(* IEC 61131-3 sources: s7-to-codesys/tests/POUs/ScenariosLang/FB_BackwashGraph_ScenarioTest, 7 files *)

(* ---- FB_BackwashGraph_ScenarioTest.decl.st ---- *)
// AUTO-GENERATED — не редактировать: s7conv gen-tests, сценарии scenarios/lang/FB_BackwashGraph.csv
// Правка — в CSV (scenarios/README.md), затем python -m s7conv build-corpus.
// Назначение: тесты поведения сконвертированного FB_BackwashGraph по сценариям CSV (сценариев: 6, строк: 46):
//             один метод-тест на сценарий, строки — по порядку с моделируемым временем GVL_S7Clock.
//             Ожидаемые значения — из CSV (эталонные модели по описанию логики блока), не из
//             результата конвертации.
// Автор:      s7conv 0.1.0 (сгенерировано)
// Версия:     не указана
// Документ:   scenarios/README.md, docs/methodology.md, раздел «Проверка поведения»
FUNCTION_BLOCK FB_BackwashGraph_ScenarioTest EXTENDS coUnit.FB_TestSuite
VAR
    fbLongWash : FB_BackwashGraph;  // свой экземпляр на сценарий
    xLongWashDone : BOOL;  // сценарий выполнен (выполняется один раз)
    fbShortWash : FB_BackwashGraph;  // свой экземпляр на сценарий
    xShortWashDone : BOOL;  // сценарий выполнен (выполняется один раз)
    fbSupervision : FB_BackwashGraph;  // свой экземпляр на сценарий
    xSupervisionDone : BOOL;  // сценарий выполнен (выполняется один раз)
    fbAckSwitches : FB_BackwashGraph;  // свой экземпляр на сценарий
    xAckSwitchesDone : BOOL;  // сценарий выполнен (выполняется один раз)
    fbInterlockPump : FB_BackwashGraph;  // свой экземпляр на сценарий
    xInterlockPumpDone : BOOL;  // сценарий выполнен (выполняется один раз)
    fbOffAndInit : FB_BackwashGraph;  // свой экземпляр на сценарий
    xOffAndInitDone : BOOL;  // сценарий выполнен (выполняется один раз)
END_VAR

(* ---- AckSwitches.method.impl.st ---- *)
// AUTO-GENERATED — не редактировать: scenarios/lang/FB_BackwashGraph.csv, сценарий AckSwitches
coUnit.TEST('AckSwitches');
IF NOT xAckSwitchesDone THEN
    xAckSwitchesDone := TRUE;
    GVL_S7Clock.xSimulation := TRUE;

    // #1, t = 0 мс — первый вызов: начальный шаг Idle
    GVL_S7Clock.tSimNow := T#0MS;
    fbAckSwitches.OFF_SQ := FALSE;
    fbAckSwitches.INIT_SQ := FALSE;
    fbAckSwitches.ACK_EF := FALSE;
    fbAckSwitches.xStart := FALSE;
    fbAckSwitches.xLevelLow := FALSE;
    fbAckSwitches.xLevelHigh := FALSE;
    fbAckSwitches.xShortWash := FALSE;
    fbAckSwitches.xPumpOk := TRUE;
    fbAckSwitches.xValveFault := FALSE;
    fbAckSwitches();
    AssertEquals_BOOL(Expected := FALSE, Actual := fbAckSwitches.ERR_FLT, Message := 'AckSwitches#1 ERR_FLT');
    AssertEquals_BOOL(Expected := TRUE, Actual := fbAckSwitches.xReady, Message := 'AckSwitches#1 xReady');
    AssertEquals_BOOL(Expected := FALSE, Actual := fbAckSwitches.xDrainValve, Message := 'AckSwitches#1 xDrainValve');
    AssertEquals_BOOL(Expected := FALSE, Actual := fbAckSwitches.xBlower, Message := 'AckSwitches#1 xBlower');
    AssertEquals_BOOL(Expected := FALSE, Actual := fbAckSwitches.xAirValve, Message := 'AckSwitches#1 xAirValve');
    AssertEquals_BOOL(Expected := FALSE, Actual := fbAckSwitches.xWashPump, Message := 'AckSwitches#1 xWashPump');
    AssertEquals_BOOL(Expected := FALSE, Actual := fbAckSwitches.xInletValve, Message := 'AckSwitches#1 xInletValve');
    AssertEquals_BOOL(Expected := FALSE, Actual := fbAckSwitches.xWashActive, Message := 'AckSwitches#1 xWashActive');
    AssertEquals_BOOL(Expected := FALSE, Actual := fbAckSwitches.xValvesBusy, Message := 'AckSwitches#1 xValvesBusy');
    AssertEquals_INT(Expected := 0, Actual := fbAckSwitches.iWashCount, Message := 'AckSwitches#1 iWashCount');

    // #2, t = 100 мс — T1 Start: Drain, промывка №1, слив открыт
    GVL_S7Clock.tSimNow := T#100MS;
    fbAckSwitches.xStart := TRUE;
    fbAckSwitches();
    AssertEquals_BOOL(Expected := FALSE, Actual := fbAckSwitches.ERR_FLT, Message := 'AckSwitches#2 ERR_FLT');
    AssertEquals_BOOL(Expected := FALSE, Actual := fbAckSwitches.xReady, Message := 'AckSwitches#2 xReady');
    AssertEquals_BOOL(Expected := TRUE, Actual := fbAckSwitches.xDrainValve, Message := 'AckSwitches#2 xDrainValve');
    AssertEquals_BOOL(Expected := FALSE, Actual := fbAckSwitches.xBlower, Message := 'AckSwitches#2 xBlower');
    AssertEquals_BOOL(Expected := FALSE, Actual := fbAckSwitches.xAirValve, Message := 'AckSwitches#2 xAirValve');
    AssertEquals_BOOL(Expected := FALSE, Actual := fbAckSwitches.xWashPump, Message := 'AckSwitches#2 xWashPump');
    AssertEquals_BOOL(Expected := FALSE, Actual := fbAckSwitches.xInletValve, Message := 'AckSwitches#2 xInletValve');
    AssertEquals_BOOL(Expected := TRUE, Actual := fbAckSwitches.xWashActive, Message := 'AckSwitches#2 xWashActive');
    AssertEquals_BOOL(Expected := TRUE, Actual := fbAckSwitches.xValvesBusy, Message := 'AckSwitches#2 xValvesBusy');
    AssertEquals_INT(Expected := 1, Actual := fbAckSwitches.iWashCount, Message := 'AckSwitches#2 iWashCount');

    // #3, t = 200 мс — слив
    GVL_S7Clock.tSimNow := T#200MS;
    fbAckSwitches.xStart := FALSE;
    fbAckSwitches();
    AssertEquals_BOOL(Expected := FALSE, Actual := fbAckSwitches.ERR_FLT, Message := 'AckSwitches#3 ERR_FLT');
    AssertEquals_BOOL(Expected := FALSE, Actual := fbAckSwitches.xReady, Message := 'AckSwitches#3 xReady');
    AssertEquals_BOOL(Expected := TRUE, Actual := fbAckSwitches.xDrainValve, Message := 'AckSwitches#3 xDrainValve');
    AssertEquals_BOOL(Expected := FALSE, Actual := fbAckSwitches.xBlower, Message := 'AckSwitches#3 xBlower');
    AssertEquals_BOOL(Expected := FALSE, Actual := fbAckSwitches.xAirValve, Message := 'AckSwitches#3 xAirValve');
    AssertEquals_BOOL(Expected := FALSE, Actual := fbAckSwitches.xWashPump, Message := 'AckSwitches#3 xWashPump');
    AssertEquals_BOOL(Expected := FALSE, Actual := fbAckSwitches.xInletValve, Message := 'AckSwitches#3 xInletValve');
    AssertEquals_BOOL(Expected := TRUE, Actual := fbAckSwitches.xWashActive, Message := 'AckSwitches#3 xWashActive');
    AssertEquals_BOOL(Expected := TRUE, Actual := fbAckSwitches.xValvesBusy, Message := 'AckSwitches#3 xValvesBusy');
    AssertEquals_INT(Expected := 1, Actual := fbAckSwitches.iWashCount, Message := 'AckSwitches#3 iWashCount');

    // #4, t = 500 мс — ошибка контроля
    GVL_S7Clock.tSimNow := T#500MS;
    fbAckSwitches.xShortWash := TRUE;
    fbAckSwitches.xValveFault := TRUE;
    fbAckSwitches();
    AssertEquals_BOOL(Expected := TRUE, Actual := fbAckSwitches.ERR_FLT, Message := 'AckSwitches#4 ERR_FLT');
    AssertEquals_BOOL(Expected := FALSE, Actual := fbAckSwitches.xReady, Message := 'AckSwitches#4 xReady');
    AssertEquals_BOOL(Expected := TRUE, Actual := fbAckSwitches.xDrainValve, Message := 'AckSwitches#4 xDrainValve');
    AssertEquals_BOOL(Expected := FALSE, Actual := fbAckSwitches.xBlower, Message := 'AckSwitches#4 xBlower');
    AssertEquals_BOOL(Expected := FALSE, Actual := fbAckSwitches.xAirValve, Message := 'AckSwitches#4 xAirValve');
    AssertEquals_BOOL(Expected := FALSE, Actual := fbAckSwitches.xWashPump, Message := 'AckSwitches#4 xWashPump');
    AssertEquals_BOOL(Expected := FALSE, Actual := fbAckSwitches.xInletValve, Message := 'AckSwitches#4 xInletValve');
    AssertEquals_BOOL(Expected := TRUE, Actual := fbAckSwitches.xWashActive, Message := 'AckSwitches#4 xWashActive');
    AssertEquals_BOOL(Expected := TRUE, Actual := fbAckSwitches.xValvesBusy, Message := 'AckSwitches#4 xValvesBusy');
    AssertEquals_INT(Expected := 1, Actual := fbAckSwitches.iWashCount, Message := 'AckSwitches#4 iWashCount');

    // #5, t = 600 мс — квитирование и уровень: T3 ShortWash в том же вызове
    GVL_S7Clock.tSimNow := T#600MS;
    fbAckSwitches.ACK_EF := TRUE;
    fbAckSwitches.xLevelLow := TRUE;
    fbAckSwitches();
    AssertEquals_BOOL(Expected := FALSE, Actual := fbAckSwitches.ERR_FLT, Message := 'AckSwitches#5 ERR_FLT');
    AssertEquals_BOOL(Expected := FALSE, Actual := fbAckSwitches.xReady, Message := 'AckSwitches#5 xReady');
    AssertEquals_BOOL(Expected := FALSE, Actual := fbAckSwitches.xDrainValve, Message := 'AckSwitches#5 xDrainValve');
    AssertEquals_BOOL(Expected := FALSE, Actual := fbAckSwitches.xBlower, Message := 'AckSwitches#5 xBlower');
    AssertEquals_BOOL(Expected := FALSE, Actual := fbAckSwitches.xAirValve, Message := 'AckSwitches#5 xAirValve');
    AssertEquals_BOOL(Expected := TRUE, Actual := fbAckSwitches.xWashPump, Message := 'AckSwitches#5 xWashPump');
    AssertEquals_BOOL(Expected := FALSE, Actual := fbAckSwitches.xInletValve, Message := 'AckSwitches#5 xInletValve');
    AssertEquals_BOOL(Expected := TRUE, Actual := fbAckSwitches.xWashActive, Message := 'AckSwitches#5 xWashActive');
    AssertEquals_BOOL(Expected := FALSE, Actual := fbAckSwitches.xValvesBusy, Message := 'AckSwitches#5 xValvesBusy');
    AssertEquals_INT(Expected := 1, Actual := fbAckSwitches.iWashCount, Message := 'AckSwitches#5 iWashCount');

    // #6, t = 700 мс — QuickRinse: контроль Drain больше не действует
    GVL_S7Clock.tSimNow := T#700MS;
    fbAckSwitches.ACK_EF := FALSE;
    fbAckSwitches.xLevelLow := FALSE;
    fbAckSwitches();
    AssertEquals_BOOL(Expected := FALSE, Actual := fbAckSwitches.ERR_FLT, Message := 'AckSwitches#6 ERR_FLT');
    AssertEquals_BOOL(Expected := FALSE, Actual := fbAckSwitches.xReady, Message := 'AckSwitches#6 xReady');
    AssertEquals_BOOL(Expected := FALSE, Actual := fbAckSwitches.xDrainValve, Message := 'AckSwitches#6 xDrainValve');
    AssertEquals_BOOL(Expected := FALSE, Actual := fbAckSwitches.xBlower, Message := 'AckSwitches#6 xBlower');
    AssertEquals_BOOL(Expected := FALSE, Actual := fbAckSwitches.xAirValve, Message := 'AckSwitches#6 xAirValve');
    AssertEquals_BOOL(Expected := TRUE, Actual := fbAckSwitches.xWashPump, Message := 'AckSwitches#6 xWashPump');
    AssertEquals_BOOL(Expected := FALSE, Actual := fbAckSwitches.xInletValve, Message := 'AckSwitches#6 xInletValve');
    AssertEquals_BOOL(Expected := TRUE, Actual := fbAckSwitches.xWashActive, Message := 'AckSwitches#6 xWashActive');
    AssertEquals_BOOL(Expected := FALSE, Actual := fbAckSwitches.xValvesBusy, Message := 'AckSwitches#6 xValvesBusy');
    AssertEquals_INT(Expected := 1, Actual := fbAckSwitches.iWashCount, Message := 'AckSwitches#6 iWashCount');

    GVL_S7Clock.xSimulation := FALSE;
END_IF
coUnit.TEST_FINISHED();

(* ---- InterlockPump.method.impl.st ---- *)
// AUTO-GENERATED — не редактировать: scenarios/lang/FB_BackwashGraph.csv, сценарий InterlockPump
coUnit.TEST('InterlockPump');
IF NOT xInterlockPumpDone THEN
    xInterlockPumpDone := TRUE;
    GVL_S7Clock.xSimulation := TRUE;

    // #1, t = 0 мс — первый вызов: начальный шаг Idle
    GVL_S7Clock.tSimNow := T#0MS;
    fbInterlockPump.OFF_SQ := FALSE;
    fbInterlockPump.INIT_SQ := FALSE;
    fbInterlockPump.ACK_EF := FALSE;
    fbInterlockPump.xStart := FALSE;
    fbInterlockPump.xLevelLow := FALSE;
    fbInterlockPump.xLevelHigh := FALSE;
    fbInterlockPump.xShortWash := FALSE;
    fbInterlockPump.xPumpOk := TRUE;
    fbInterlockPump.xValveFault := FALSE;
    fbInterlockPump();
    AssertEquals_BOOL(Expected := FALSE, Actual := fbInterlockPump.ERR_FLT, Message := 'InterlockPump#1 ERR_FLT');
    AssertEquals_BOOL(Expected := TRUE, Actual := fbInterlockPump.xReady, Message := 'InterlockPump#1 xReady');
    AssertEquals_BOOL(Expected := FALSE,
                      Actual := fbInterlockPump.xDrainValve,
                      Message := 'InterlockPump#1 xDrainValve');
    AssertEquals_BOOL(Expected := FALSE, Actual := fbInterlockPump.xBlower, Message := 'InterlockPump#1 xBlower');
    AssertEquals_BOOL(Expected := FALSE, Actual := fbInterlockPump.xAirValve, Message := 'InterlockPump#1 xAirValve');
    AssertEquals_BOOL(Expected := FALSE, Actual := fbInterlockPump.xWashPump, Message := 'InterlockPump#1 xWashPump');
    AssertEquals_BOOL(Expected := FALSE,
                      Actual := fbInterlockPump.xInletValve,
                      Message := 'InterlockPump#1 xInletValve');
    AssertEquals_BOOL(Expected := FALSE,
                      Actual := fbInterlockPump.xWashActive,
                      Message := 'InterlockPump#1 xWashActive');
    AssertEquals_BOOL(Expected := FALSE,
                      Actual := fbInterlockPump.xValvesBusy,
                      Message := 'InterlockPump#1 xValvesBusy');
    AssertEquals_INT(Expected := 0, Actual := fbInterlockPump.iWashCount, Message := 'InterlockPump#1 iWashCount');

    // #2, t = 100 мс — T1 Start: Drain, промывка №1, слив открыт
    GVL_S7Clock.tSimNow := T#100MS;
    fbInterlockPump.xStart := TRUE;
    fbInterlockPump();
    AssertEquals_BOOL(Expected := FALSE, Actual := fbInterlockPump.ERR_FLT, Message := 'InterlockPump#2 ERR_FLT');
    AssertEquals_BOOL(Expected := FALSE, Actual := fbInterlockPump.xReady, Message := 'InterlockPump#2 xReady');
    AssertEquals_BOOL(Expected := TRUE,
                      Actual := fbInterlockPump.xDrainValve,
                      Message := 'InterlockPump#2 xDrainValve');
    AssertEquals_BOOL(Expected := FALSE, Actual := fbInterlockPump.xBlower, Message := 'InterlockPump#2 xBlower');
    AssertEquals_BOOL(Expected := FALSE, Actual := fbInterlockPump.xAirValve, Message := 'InterlockPump#2 xAirValve');
    AssertEquals_BOOL(Expected := FALSE, Actual := fbInterlockPump.xWashPump, Message := 'InterlockPump#2 xWashPump');
    AssertEquals_BOOL(Expected := FALSE,
                      Actual := fbInterlockPump.xInletValve,
                      Message := 'InterlockPump#2 xInletValve');
    AssertEquals_BOOL(Expected := TRUE,
                      Actual := fbInterlockPump.xWashActive,
                      Message := 'InterlockPump#2 xWashActive');
    AssertEquals_BOOL(Expected := TRUE,
                      Actual := fbInterlockPump.xValvesBusy,
                      Message := 'InterlockPump#2 xValvesBusy');
    AssertEquals_INT(Expected := 1, Actual := fbInterlockPump.iWashCount, Message := 'InterlockPump#2 iWashCount');

    // #3, t = 200 мс — слив
    GVL_S7Clock.tSimNow := T#200MS;
    fbInterlockPump.xStart := FALSE;
    fbInterlockPump();
    AssertEquals_BOOL(Expected := FALSE, Actual := fbInterlockPump.ERR_FLT, Message := 'InterlockPump#3 ERR_FLT');
    AssertEquals_BOOL(Expected := FALSE, Actual := fbInterlockPump.xReady, Message := 'InterlockPump#3 xReady');
    AssertEquals_BOOL(Expected := TRUE,
                      Actual := fbInterlockPump.xDrainValve,
                      Message := 'InterlockPump#3 xDrainValve');
    AssertEquals_BOOL(Expected := FALSE, Actual := fbInterlockPump.xBlower, Message := 'InterlockPump#3 xBlower');
    AssertEquals_BOOL(Expected := FALSE, Actual := fbInterlockPump.xAirValve, Message := 'InterlockPump#3 xAirValve');
    AssertEquals_BOOL(Expected := FALSE, Actual := fbInterlockPump.xWashPump, Message := 'InterlockPump#3 xWashPump');
    AssertEquals_BOOL(Expected := FALSE,
                      Actual := fbInterlockPump.xInletValve,
                      Message := 'InterlockPump#3 xInletValve');
    AssertEquals_BOOL(Expected := TRUE,
                      Actual := fbInterlockPump.xWashActive,
                      Message := 'InterlockPump#3 xWashActive');
    AssertEquals_BOOL(Expected := TRUE,
                      Actual := fbInterlockPump.xValvesBusy,
                      Message := 'InterlockPump#3 xValvesBusy');
    AssertEquals_INT(Expected := 1, Actual := fbInterlockPump.iWashCount, Message := 'InterlockPump#3 iWashCount');

    // #4, t = 1000 мс — Air и Rinse: насос промывки включён
    GVL_S7Clock.tSimNow := T#1000MS;
    fbInterlockPump.xLevelLow := TRUE;
    fbInterlockPump();
    AssertEquals_BOOL(Expected := FALSE, Actual := fbInterlockPump.ERR_FLT, Message := 'InterlockPump#4 ERR_FLT');
    AssertEquals_BOOL(Expected := FALSE, Actual := fbInterlockPump.xReady, Message := 'InterlockPump#4 xReady');
    AssertEquals_BOOL(Expected := FALSE,
                      Actual := fbInterlockPump.xDrainValve,
                      Message := 'InterlockPump#4 xDrainValve');
    AssertEquals_BOOL(Expected := TRUE, Actual := fbInterlockPump.xBlower, Message := 'InterlockPump#4 xBlower');
    AssertEquals_BOOL(Expected := FALSE, Actual := fbInterlockPump.xAirValve, Message := 'InterlockPump#4 xAirValve');
    AssertEquals_BOOL(Expected := TRUE, Actual := fbInterlockPump.xWashPump, Message := 'InterlockPump#4 xWashPump');
    AssertEquals_BOOL(Expected := FALSE,
                      Actual := fbInterlockPump.xInletValve,
                      Message := 'InterlockPump#4 xInletValve');
    AssertEquals_BOOL(Expected := TRUE,
                      Actual := fbInterlockPump.xWashActive,
                      Message := 'InterlockPump#4 xWashActive');
    AssertEquals_BOOL(Expected := FALSE,
                      Actual := fbInterlockPump.xValvesBusy,
                      Message := 'InterlockPump#4 xValvesBusy');
    AssertEquals_INT(Expected := 1, Actual := fbInterlockPump.iWashCount, Message := 'InterlockPump#4 iWashCount');

    // #5, t = 1100 мс — насос неисправен: блокировка не выполнена
    GVL_S7Clock.tSimNow := T#1100MS;
    fbInterlockPump.xLevelLow := FALSE;
    fbInterlockPump.xPumpOk := FALSE;
    fbInterlockPump();
    AssertEquals_BOOL(Expected := FALSE, Actual := fbInterlockPump.ERR_FLT, Message := 'InterlockPump#5 ERR_FLT');
    AssertEquals_BOOL(Expected := FALSE, Actual := fbInterlockPump.xReady, Message := 'InterlockPump#5 xReady');
    AssertEquals_BOOL(Expected := FALSE,
                      Actual := fbInterlockPump.xDrainValve,
                      Message := 'InterlockPump#5 xDrainValve');
    AssertEquals_BOOL(Expected := TRUE, Actual := fbInterlockPump.xBlower, Message := 'InterlockPump#5 xBlower');
    AssertEquals_BOOL(Expected := FALSE, Actual := fbInterlockPump.xAirValve, Message := 'InterlockPump#5 xAirValve');
    AssertEquals_BOOL(Expected := FALSE, Actual := fbInterlockPump.xWashPump, Message := 'InterlockPump#5 xWashPump');
    AssertEquals_BOOL(Expected := FALSE,
                      Actual := fbInterlockPump.xInletValve,
                      Message := 'InterlockPump#5 xInletValve');
    AssertEquals_BOOL(Expected := TRUE,
                      Actual := fbInterlockPump.xWashActive,
                      Message := 'InterlockPump#5 xWashActive');
    AssertEquals_BOOL(Expected := FALSE,
                      Actual := fbInterlockPump.xValvesBusy,
                      Message := 'InterlockPump#5 xValvesBusy');
    AssertEquals_INT(Expected := 1, Actual := fbInterlockPump.iWashCount, Message := 'InterlockPump#5 iWashCount');

    // #6, t = 1200 мс — насос исправен: снова включён
    GVL_S7Clock.tSimNow := T#1200MS;
    fbInterlockPump.xPumpOk := TRUE;
    fbInterlockPump();
    AssertEquals_BOOL(Expected := FALSE, Actual := fbInterlockPump.ERR_FLT, Message := 'InterlockPump#6 ERR_FLT');
    AssertEquals_BOOL(Expected := FALSE, Actual := fbInterlockPump.xReady, Message := 'InterlockPump#6 xReady');
    AssertEquals_BOOL(Expected := FALSE,
                      Actual := fbInterlockPump.xDrainValve,
                      Message := 'InterlockPump#6 xDrainValve');
    AssertEquals_BOOL(Expected := TRUE, Actual := fbInterlockPump.xBlower, Message := 'InterlockPump#6 xBlower');
    AssertEquals_BOOL(Expected := FALSE, Actual := fbInterlockPump.xAirValve, Message := 'InterlockPump#6 xAirValve');
    AssertEquals_BOOL(Expected := TRUE, Actual := fbInterlockPump.xWashPump, Message := 'InterlockPump#6 xWashPump');
    AssertEquals_BOOL(Expected := FALSE,
                      Actual := fbInterlockPump.xInletValve,
                      Message := 'InterlockPump#6 xInletValve');
    AssertEquals_BOOL(Expected := TRUE,
                      Actual := fbInterlockPump.xWashActive,
                      Message := 'InterlockPump#6 xWashActive');
    AssertEquals_BOOL(Expected := FALSE,
                      Actual := fbInterlockPump.xValvesBusy,
                      Message := 'InterlockPump#6 xValvesBusy');
    AssertEquals_INT(Expected := 1, Actual := fbInterlockPump.iWashCount, Message := 'InterlockPump#6 iWashCount');

    GVL_S7Clock.xSimulation := FALSE;
END_IF
coUnit.TEST_FINISHED();

(* ---- LongWash.method.impl.st ---- *)
// AUTO-GENERATED — не редактировать: scenarios/lang/FB_BackwashGraph.csv, сценарий LongWash
coUnit.TEST('LongWash');
IF NOT xLongWashDone THEN
    xLongWashDone := TRUE;
    GVL_S7Clock.xSimulation := TRUE;

    // #1, t = 0 мс — первый вызов: начальный шаг Idle
    GVL_S7Clock.tSimNow := T#0MS;
    fbLongWash.OFF_SQ := FALSE;
    fbLongWash.INIT_SQ := FALSE;
    fbLongWash.ACK_EF := FALSE;
    fbLongWash.xStart := FALSE;
    fbLongWash.xLevelLow := FALSE;
    fbLongWash.xLevelHigh := FALSE;
    fbLongWash.xShortWash := FALSE;
    fbLongWash.xPumpOk := TRUE;
    fbLongWash.xValveFault := FALSE;
    fbLongWash();
    AssertEquals_BOOL(Expected := FALSE, Actual := fbLongWash.ERR_FLT, Message := 'LongWash#1 ERR_FLT');
    AssertEquals_BOOL(Expected := TRUE, Actual := fbLongWash.xReady, Message := 'LongWash#1 xReady');
    AssertEquals_BOOL(Expected := FALSE, Actual := fbLongWash.xDrainValve, Message := 'LongWash#1 xDrainValve');
    AssertEquals_BOOL(Expected := FALSE, Actual := fbLongWash.xBlower, Message := 'LongWash#1 xBlower');
    AssertEquals_BOOL(Expected := FALSE, Actual := fbLongWash.xAirValve, Message := 'LongWash#1 xAirValve');
    AssertEquals_BOOL(Expected := FALSE, Actual := fbLongWash.xWashPump, Message := 'LongWash#1 xWashPump');
    AssertEquals_BOOL(Expected := FALSE, Actual := fbLongWash.xInletValve, Message := 'LongWash#1 xInletValve');
    AssertEquals_BOOL(Expected := FALSE, Actual := fbLongWash.xWashActive, Message := 'LongWash#1 xWashActive');
    AssertEquals_BOOL(Expected := FALSE, Actual := fbLongWash.xValvesBusy, Message := 'LongWash#1 xValvesBusy');
    AssertEquals_INT(Expected := 0, Actual := fbLongWash.iWashCount, Message := 'LongWash#1 iWashCount');

    // #2, t = 100 мс — T1 Start: Drain, промывка №1, слив открыт
    GVL_S7Clock.tSimNow := T#100MS;
    fbLongWash.xStart := TRUE;
    fbLongWash();
    AssertEquals_BOOL(Expected := FALSE, Actual := fbLongWash.ERR_FLT, Message := 'LongWash#2 ERR_FLT');
    AssertEquals_BOOL(Expected := FALSE, Actual := fbLongWash.xReady, Message := 'LongWash#2 xReady');
    AssertEquals_BOOL(Expected := TRUE, Actual := fbLongWash.xDrainValve, Message := 'LongWash#2 xDrainValve');
    AssertEquals_BOOL(Expected := FALSE, Actual := fbLongWash.xBlower, Message := 'LongWash#2 xBlower');
    AssertEquals_BOOL(Expected := FALSE, Actual := fbLongWash.xAirValve, Message := 'LongWash#2 xAirValve');
    AssertEquals_BOOL(Expected := FALSE, Actual := fbLongWash.xWashPump, Message := 'LongWash#2 xWashPump');
    AssertEquals_BOOL(Expected := FALSE, Actual := fbLongWash.xInletValve, Message := 'LongWash#2 xInletValve');
    AssertEquals_BOOL(Expected := TRUE, Actual := fbLongWash.xWashActive, Message := 'LongWash#2 xWashActive');
    AssertEquals_BOOL(Expected := TRUE, Actual := fbLongWash.xValvesBusy, Message := 'LongWash#2 xValvesBusy');
    AssertEquals_INT(Expected := 1, Actual := fbLongWash.iWashCount, Message := 'LongWash#2 iWashCount');

    // #3, t = 200 мс — слив
    GVL_S7Clock.tSimNow := T#200MS;
    fbLongWash.xStart := FALSE;
    fbLongWash();
    AssertEquals_BOOL(Expected := FALSE, Actual := fbLongWash.ERR_FLT, Message := 'LongWash#3 ERR_FLT');
    AssertEquals_BOOL(Expected := FALSE, Actual := fbLongWash.xReady, Message := 'LongWash#3 xReady');
    AssertEquals_BOOL(Expected := TRUE, Actual := fbLongWash.xDrainValve, Message := 'LongWash#3 xDrainValve');
    AssertEquals_BOOL(Expected := FALSE, Actual := fbLongWash.xBlower, Message := 'LongWash#3 xBlower');
    AssertEquals_BOOL(Expected := FALSE, Actual := fbLongWash.xAirValve, Message := 'LongWash#3 xAirValve');
    AssertEquals_BOOL(Expected := FALSE, Actual := fbLongWash.xWashPump, Message := 'LongWash#3 xWashPump');
    AssertEquals_BOOL(Expected := FALSE, Actual := fbLongWash.xInletValve, Message := 'LongWash#3 xInletValve');
    AssertEquals_BOOL(Expected := TRUE, Actual := fbLongWash.xWashActive, Message := 'LongWash#3 xWashActive');
    AssertEquals_BOOL(Expected := TRUE, Actual := fbLongWash.xValvesBusy, Message := 'LongWash#3 xValvesBusy');
    AssertEquals_INT(Expected := 1, Actual := fbLongWash.iWashCount, Message := 'LongWash#3 iWashCount');

    // #4, t = 1000 мс — T2 LongWash: параллельно Air и Rinse
    GVL_S7Clock.tSimNow := T#1000MS;
    fbLongWash.xLevelLow := TRUE;
    fbLongWash();
    AssertEquals_BOOL(Expected := FALSE, Actual := fbLongWash.ERR_FLT, Message := 'LongWash#4 ERR_FLT');
    AssertEquals_BOOL(Expected := FALSE, Actual := fbLongWash.xReady, Message := 'LongWash#4 xReady');
    AssertEquals_BOOL(Expected := FALSE, Actual := fbLongWash.xDrainValve, Message := 'LongWash#4 xDrainValve');
    AssertEquals_BOOL(Expected := TRUE, Actual := fbLongWash.xBlower, Message := 'LongWash#4 xBlower');
    AssertEquals_BOOL(Expected := FALSE, Actual := fbLongWash.xAirValve, Message := 'LongWash#4 xAirValve');
    AssertEquals_BOOL(Expected := TRUE, Actual := fbLongWash.xWashPump, Message := 'LongWash#4 xWashPump');
    AssertEquals_BOOL(Expected := FALSE, Actual := fbLongWash.xInletValve, Message := 'LongWash#4 xInletValve');
    AssertEquals_BOOL(Expected := TRUE, Actual := fbLongWash.xWashActive, Message := 'LongWash#4 xWashActive');
    AssertEquals_BOOL(Expected := FALSE, Actual := fbLongWash.xValvesBusy, Message := 'LongWash#4 xValvesBusy');
    AssertEquals_INT(Expected := 1, Actual := fbLongWash.iWashCount, Message := 'LongWash#4 iWashCount');

    // #5, t = 1100 мс — воздуходувка и насос; задвижка воздуха ещё закрыта
    GVL_S7Clock.tSimNow := T#1100MS;
    fbLongWash.xLevelLow := FALSE;
    fbLongWash();
    AssertEquals_BOOL(Expected := FALSE, Actual := fbLongWash.ERR_FLT, Message := 'LongWash#5 ERR_FLT');
    AssertEquals_BOOL(Expected := FALSE, Actual := fbLongWash.xReady, Message := 'LongWash#5 xReady');
    AssertEquals_BOOL(Expected := FALSE, Actual := fbLongWash.xDrainValve, Message := 'LongWash#5 xDrainValve');
    AssertEquals_BOOL(Expected := TRUE, Actual := fbLongWash.xBlower, Message := 'LongWash#5 xBlower');
    AssertEquals_BOOL(Expected := FALSE, Actual := fbLongWash.xAirValve, Message := 'LongWash#5 xAirValve');
    AssertEquals_BOOL(Expected := TRUE, Actual := fbLongWash.xWashPump, Message := 'LongWash#5 xWashPump');
    AssertEquals_BOOL(Expected := FALSE, Actual := fbLongWash.xInletValve, Message := 'LongWash#5 xInletValve');
    AssertEquals_BOOL(Expected := TRUE, Actual := fbLongWash.xWashActive, Message := 'LongWash#5 xWashActive');
    AssertEquals_BOOL(Expected := FALSE, Actual := fbLongWash.xValvesBusy, Message := 'LongWash#5 xValvesBusy');
    AssertEquals_INT(Expected := 1, Actual := fbLongWash.iWashCount, Message := 'LongWash#5 iWashCount');

    // #6, t = 3000 мс, на пороге таймера — 2 с продувки: задвижка воздуха открыта (D)
    GVL_S7Clock.tSimNow := T#3000MS;
    fbLongWash();
    AssertEquals_BOOL(Expected := FALSE, Actual := fbLongWash.ERR_FLT, Message := 'LongWash#6 ERR_FLT');
    AssertEquals_BOOL(Expected := FALSE, Actual := fbLongWash.xReady, Message := 'LongWash#6 xReady');
    AssertEquals_BOOL(Expected := FALSE, Actual := fbLongWash.xDrainValve, Message := 'LongWash#6 xDrainValve');
    AssertEquals_BOOL(Expected := TRUE, Actual := fbLongWash.xBlower, Message := 'LongWash#6 xBlower');
    AssertEquals_BOOL(Expected := TRUE, Actual := fbLongWash.xAirValve, Message := 'LongWash#6 xAirValve');
    AssertEquals_BOOL(Expected := TRUE, Actual := fbLongWash.xWashPump, Message := 'LongWash#6 xWashPump');
    AssertEquals_BOOL(Expected := FALSE, Actual := fbLongWash.xInletValve, Message := 'LongWash#6 xInletValve');
    AssertEquals_BOOL(Expected := TRUE, Actual := fbLongWash.xWashActive, Message := 'LongWash#6 xWashActive');
    AssertEquals_BOOL(Expected := FALSE, Actual := fbLongWash.xValvesBusy, Message := 'LongWash#6 xValvesBusy');
    AssertEquals_INT(Expected := 1, Actual := fbLongWash.iWashCount, Message := 'LongWash#6 iWashCount');

    // #7, t = 10700 мс — 9,7 с: синхронизация ещё не прошла
    GVL_S7Clock.tSimNow := T#10700MS;
    fbLongWash();
    AssertEquals_BOOL(Expected := FALSE, Actual := fbLongWash.ERR_FLT, Message := 'LongWash#7 ERR_FLT');
    AssertEquals_BOOL(Expected := FALSE, Actual := fbLongWash.xReady, Message := 'LongWash#7 xReady');
    AssertEquals_BOOL(Expected := FALSE, Actual := fbLongWash.xDrainValve, Message := 'LongWash#7 xDrainValve');
    AssertEquals_BOOL(Expected := TRUE, Actual := fbLongWash.xBlower, Message := 'LongWash#7 xBlower');
    AssertEquals_BOOL(Expected := TRUE, Actual := fbLongWash.xAirValve, Message := 'LongWash#7 xAirValve');
    AssertEquals_BOOL(Expected := TRUE, Actual := fbLongWash.xWashPump, Message := 'LongWash#7 xWashPump');
    AssertEquals_BOOL(Expected := FALSE, Actual := fbLongWash.xInletValve, Message := 'LongWash#7 xInletValve');
    AssertEquals_BOOL(Expected := TRUE, Actual := fbLongWash.xWashActive, Message := 'LongWash#7 xWashActive');
    AssertEquals_BOOL(Expected := FALSE, Actual := fbLongWash.xValvesBusy, Message := 'LongWash#7 xValvesBusy');
    AssertEquals_INT(Expected := 1, Actual := fbLongWash.iWashCount, Message := 'LongWash#7 iWashCount');

    // #8, t = 11000 мс, на пороге таймера — 10 с: T4 AirDone — Refill, подача открыта
    GVL_S7Clock.tSimNow := T#11000MS;
    fbLongWash();
    AssertEquals_BOOL(Expected := FALSE, Actual := fbLongWash.ERR_FLT, Message := 'LongWash#8 ERR_FLT');
    AssertEquals_BOOL(Expected := FALSE, Actual := fbLongWash.xReady, Message := 'LongWash#8 xReady');
    AssertEquals_BOOL(Expected := FALSE, Actual := fbLongWash.xDrainValve, Message := 'LongWash#8 xDrainValve');
    AssertEquals_BOOL(Expected := FALSE, Actual := fbLongWash.xBlower, Message := 'LongWash#8 xBlower');
    AssertEquals_BOOL(Expected := FALSE, Actual := fbLongWash.xAirValve, Message := 'LongWash#8 xAirValve');
    AssertEquals_BOOL(Expected := FALSE, Actual := fbLongWash.xWashPump, Message := 'LongWash#8 xWashPump');
    AssertEquals_BOOL(Expected := TRUE, Actual := fbLongWash.xInletValve, Message := 'LongWash#8 xInletValve');
    AssertEquals_BOOL(Expected := FALSE, Actual := fbLongWash.xWashActive, Message := 'LongWash#8 xWashActive');
    AssertEquals_BOOL(Expected := TRUE, Actual := fbLongWash.xValvesBusy, Message := 'LongWash#8 xValvesBusy');
    AssertEquals_INT(Expected := 1, Actual := fbLongWash.iWashCount, Message := 'LongWash#8 iWashCount');

    // #9, t = 11500 мс — T6 Full: прыжок к Idle
    GVL_S7Clock.tSimNow := T#11500MS;
    fbLongWash.xLevelHigh := TRUE;
    fbLongWash();
    AssertEquals_BOOL(Expected := FALSE, Actual := fbLongWash.ERR_FLT, Message := 'LongWash#9 ERR_FLT');
    AssertEquals_BOOL(Expected := TRUE, Actual := fbLongWash.xReady, Message := 'LongWash#9 xReady');
    AssertEquals_BOOL(Expected := FALSE, Actual := fbLongWash.xDrainValve, Message := 'LongWash#9 xDrainValve');
    AssertEquals_BOOL(Expected := FALSE, Actual := fbLongWash.xBlower, Message := 'LongWash#9 xBlower');
    AssertEquals_BOOL(Expected := FALSE, Actual := fbLongWash.xAirValve, Message := 'LongWash#9 xAirValve');
    AssertEquals_BOOL(Expected := FALSE, Actual := fbLongWash.xWashPump, Message := 'LongWash#9 xWashPump');
    AssertEquals_BOOL(Expected := FALSE, Actual := fbLongWash.xInletValve, Message := 'LongWash#9 xInletValve');
    AssertEquals_BOOL(Expected := FALSE, Actual := fbLongWash.xWashActive, Message := 'LongWash#9 xWashActive');
    AssertEquals_BOOL(Expected := FALSE, Actual := fbLongWash.xValvesBusy, Message := 'LongWash#9 xValvesBusy');
    AssertEquals_INT(Expected := 1, Actual := fbLongWash.iWashCount, Message := 'LongWash#9 iWashCount');

    // #10, t = 11600 мс — готов к новой промывке
    GVL_S7Clock.tSimNow := T#11600MS;
    fbLongWash.xLevelHigh := FALSE;
    fbLongWash();
    AssertEquals_BOOL(Expected := FALSE, Actual := fbLongWash.ERR_FLT, Message := 'LongWash#10 ERR_FLT');
    AssertEquals_BOOL(Expected := TRUE, Actual := fbLongWash.xReady, Message := 'LongWash#10 xReady');
    AssertEquals_BOOL(Expected := FALSE, Actual := fbLongWash.xDrainValve, Message := 'LongWash#10 xDrainValve');
    AssertEquals_BOOL(Expected := FALSE, Actual := fbLongWash.xBlower, Message := 'LongWash#10 xBlower');
    AssertEquals_BOOL(Expected := FALSE, Actual := fbLongWash.xAirValve, Message := 'LongWash#10 xAirValve');
    AssertEquals_BOOL(Expected := FALSE, Actual := fbLongWash.xWashPump, Message := 'LongWash#10 xWashPump');
    AssertEquals_BOOL(Expected := FALSE, Actual := fbLongWash.xInletValve, Message := 'LongWash#10 xInletValve');
    AssertEquals_BOOL(Expected := FALSE, Actual := fbLongWash.xWashActive, Message := 'LongWash#10 xWashActive');
    AssertEquals_BOOL(Expected := FALSE, Actual := fbLongWash.xValvesBusy, Message := 'LongWash#10 xValvesBusy');
    AssertEquals_INT(Expected := 1, Actual := fbLongWash.iWashCount, Message := 'LongWash#10 iWashCount');

    GVL_S7Clock.xSimulation := FALSE;
END_IF
coUnit.TEST_FINISHED();

(* ---- OffAndInit.method.impl.st ---- *)
// AUTO-GENERATED — не редактировать: scenarios/lang/FB_BackwashGraph.csv, сценарий OffAndInit
coUnit.TEST('OffAndInit');
IF NOT xOffAndInitDone THEN
    xOffAndInitDone := TRUE;
    GVL_S7Clock.xSimulation := TRUE;

    // #1, t = 0 мс — первый вызов: начальный шаг Idle
    GVL_S7Clock.tSimNow := T#0MS;
    fbOffAndInit.OFF_SQ := FALSE;
    fbOffAndInit.INIT_SQ := FALSE;
    fbOffAndInit.ACK_EF := FALSE;
    fbOffAndInit.xStart := FALSE;
    fbOffAndInit.xLevelLow := FALSE;
    fbOffAndInit.xLevelHigh := FALSE;
    fbOffAndInit.xShortWash := FALSE;
    fbOffAndInit.xPumpOk := TRUE;
    fbOffAndInit.xValveFault := FALSE;
    fbOffAndInit();
    AssertEquals_BOOL(Expected := FALSE, Actual := fbOffAndInit.ERR_FLT, Message := 'OffAndInit#1 ERR_FLT');
    AssertEquals_BOOL(Expected := TRUE, Actual := fbOffAndInit.xReady, Message := 'OffAndInit#1 xReady');
    AssertEquals_BOOL(Expected := FALSE, Actual := fbOffAndInit.xDrainValve, Message := 'OffAndInit#1 xDrainValve');
    AssertEquals_BOOL(Expected := FALSE, Actual := fbOffAndInit.xBlower, Message := 'OffAndInit#1 xBlower');
    AssertEquals_BOOL(Expected := FALSE, Actual := fbOffAndInit.xAirValve, Message := 'OffAndInit#1 xAirValve');
    AssertEquals_BOOL(Expected := FALSE, Actual := fbOffAndInit.xWashPump, Message := 'OffAndInit#1 xWashPump');
    AssertEquals_BOOL(Expected := FALSE, Actual := fbOffAndInit.xInletValve, Message := 'OffAndInit#1 xInletValve');
    AssertEquals_BOOL(Expected := FALSE, Actual := fbOffAndInit.xWashActive, Message := 'OffAndInit#1 xWashActive');
    AssertEquals_BOOL(Expected := FALSE, Actual := fbOffAndInit.xValvesBusy, Message := 'OffAndInit#1 xValvesBusy');
    AssertEquals_INT(Expected := 0, Actual := fbOffAndInit.iWashCount, Message := 'OffAndInit#1 iWashCount');

    // #2, t = 100 мс — T1 Start: Drain, промывка №1, слив открыт
    GVL_S7Clock.tSimNow := T#100MS;
    fbOffAndInit.xStart := TRUE;
    fbOffAndInit();
    AssertEquals_BOOL(Expected := FALSE, Actual := fbOffAndInit.ERR_FLT, Message := 'OffAndInit#2 ERR_FLT');
    AssertEquals_BOOL(Expected := FALSE, Actual := fbOffAndInit.xReady, Message := 'OffAndInit#2 xReady');
    AssertEquals_BOOL(Expected := TRUE, Actual := fbOffAndInit.xDrainValve, Message := 'OffAndInit#2 xDrainValve');
    AssertEquals_BOOL(Expected := FALSE, Actual := fbOffAndInit.xBlower, Message := 'OffAndInit#2 xBlower');
    AssertEquals_BOOL(Expected := FALSE, Actual := fbOffAndInit.xAirValve, Message := 'OffAndInit#2 xAirValve');
    AssertEquals_BOOL(Expected := FALSE, Actual := fbOffAndInit.xWashPump, Message := 'OffAndInit#2 xWashPump');
    AssertEquals_BOOL(Expected := FALSE, Actual := fbOffAndInit.xInletValve, Message := 'OffAndInit#2 xInletValve');
    AssertEquals_BOOL(Expected := TRUE, Actual := fbOffAndInit.xWashActive, Message := 'OffAndInit#2 xWashActive');
    AssertEquals_BOOL(Expected := TRUE, Actual := fbOffAndInit.xValvesBusy, Message := 'OffAndInit#2 xValvesBusy');
    AssertEquals_INT(Expected := 1, Actual := fbOffAndInit.iWashCount, Message := 'OffAndInit#2 iWashCount');

    // #3, t = 200 мс — слив
    GVL_S7Clock.tSimNow := T#200MS;
    fbOffAndInit.xStart := FALSE;
    fbOffAndInit();
    AssertEquals_BOOL(Expected := FALSE, Actual := fbOffAndInit.ERR_FLT, Message := 'OffAndInit#3 ERR_FLT');
    AssertEquals_BOOL(Expected := FALSE, Actual := fbOffAndInit.xReady, Message := 'OffAndInit#3 xReady');
    AssertEquals_BOOL(Expected := TRUE, Actual := fbOffAndInit.xDrainValve, Message := 'OffAndInit#3 xDrainValve');
    AssertEquals_BOOL(Expected := FALSE, Actual := fbOffAndInit.xBlower, Message := 'OffAndInit#3 xBlower');
    AssertEquals_BOOL(Expected := FALSE, Actual := fbOffAndInit.xAirValve, Message := 'OffAndInit#3 xAirValve');
    AssertEquals_BOOL(Expected := FALSE, Actual := fbOffAndInit.xWashPump, Message := 'OffAndInit#3 xWashPump');
    AssertEquals_BOOL(Expected := FALSE, Actual := fbOffAndInit.xInletValve, Message := 'OffAndInit#3 xInletValve');
    AssertEquals_BOOL(Expected := TRUE, Actual := fbOffAndInit.xWashActive, Message := 'OffAndInit#3 xWashActive');
    AssertEquals_BOOL(Expected := TRUE, Actual := fbOffAndInit.xValvesBusy, Message := 'OffAndInit#3 xValvesBusy');
    AssertEquals_INT(Expected := 1, Actual := fbOffAndInit.iWashCount, Message := 'OffAndInit#3 iWashCount');

    // #4, t = 300 мс — OFF_SQ: шаг Drain выключен, слив закрыт; промывка идёт (S держится)
    GVL_S7Clock.tSimNow := T#300MS;
    fbOffAndInit.OFF_SQ := TRUE;
    fbOffAndInit();
    AssertEquals_BOOL(Expected := FALSE, Actual := fbOffAndInit.ERR_FLT, Message := 'OffAndInit#4 ERR_FLT');
    AssertEquals_BOOL(Expected := FALSE, Actual := fbOffAndInit.xReady, Message := 'OffAndInit#4 xReady');
    AssertEquals_BOOL(Expected := FALSE, Actual := fbOffAndInit.xDrainValve, Message := 'OffAndInit#4 xDrainValve');
    AssertEquals_BOOL(Expected := FALSE, Actual := fbOffAndInit.xBlower, Message := 'OffAndInit#4 xBlower');
    AssertEquals_BOOL(Expected := FALSE, Actual := fbOffAndInit.xAirValve, Message := 'OffAndInit#4 xAirValve');
    AssertEquals_BOOL(Expected := FALSE, Actual := fbOffAndInit.xWashPump, Message := 'OffAndInit#4 xWashPump');
    AssertEquals_BOOL(Expected := FALSE, Actual := fbOffAndInit.xInletValve, Message := 'OffAndInit#4 xInletValve');
    AssertEquals_BOOL(Expected := TRUE, Actual := fbOffAndInit.xWashActive, Message := 'OffAndInit#4 xWashActive');
    AssertEquals_BOOL(Expected := FALSE, Actual := fbOffAndInit.xValvesBusy, Message := 'OffAndInit#4 xValvesBusy');
    AssertEquals_INT(Expected := 1, Actual := fbOffAndInit.iWashCount, Message := 'OffAndInit#4 iWashCount');

    // #5, t = 400 мс — пуск без активных шагов: ничего
    GVL_S7Clock.tSimNow := T#400MS;
    fbOffAndInit.OFF_SQ := FALSE;
    fbOffAndInit.xStart := TRUE;
    fbOffAndInit();
    AssertEquals_BOOL(Expected := FALSE, Actual := fbOffAndInit.ERR_FLT, Message := 'OffAndInit#5 ERR_FLT');
    AssertEquals_BOOL(Expected := FALSE, Actual := fbOffAndInit.xReady, Message := 'OffAndInit#5 xReady');
    AssertEquals_BOOL(Expected := FALSE, Actual := fbOffAndInit.xDrainValve, Message := 'OffAndInit#5 xDrainValve');
    AssertEquals_BOOL(Expected := FALSE, Actual := fbOffAndInit.xBlower, Message := 'OffAndInit#5 xBlower');
    AssertEquals_BOOL(Expected := FALSE, Actual := fbOffAndInit.xAirValve, Message := 'OffAndInit#5 xAirValve');
    AssertEquals_BOOL(Expected := FALSE, Actual := fbOffAndInit.xWashPump, Message := 'OffAndInit#5 xWashPump');
    AssertEquals_BOOL(Expected := FALSE, Actual := fbOffAndInit.xInletValve, Message := 'OffAndInit#5 xInletValve');
    AssertEquals_BOOL(Expected := TRUE, Actual := fbOffAndInit.xWashActive, Message := 'OffAndInit#5 xWashActive');
    AssertEquals_BOOL(Expected := FALSE, Actual := fbOffAndInit.xValvesBusy, Message := 'OffAndInit#5 xValvesBusy');
    AssertEquals_INT(Expected := 1, Actual := fbOffAndInit.iWashCount, Message := 'OffAndInit#5 iWashCount');

    // #6, t = 500 мс — INIT_SQ: Idle
    GVL_S7Clock.tSimNow := T#500MS;
    fbOffAndInit.INIT_SQ := TRUE;
    fbOffAndInit.xStart := FALSE;
    fbOffAndInit();
    AssertEquals_BOOL(Expected := FALSE, Actual := fbOffAndInit.ERR_FLT, Message := 'OffAndInit#6 ERR_FLT');
    AssertEquals_BOOL(Expected := TRUE, Actual := fbOffAndInit.xReady, Message := 'OffAndInit#6 xReady');
    AssertEquals_BOOL(Expected := FALSE, Actual := fbOffAndInit.xDrainValve, Message := 'OffAndInit#6 xDrainValve');
    AssertEquals_BOOL(Expected := FALSE, Actual := fbOffAndInit.xBlower, Message := 'OffAndInit#6 xBlower');
    AssertEquals_BOOL(Expected := FALSE, Actual := fbOffAndInit.xAirValve, Message := 'OffAndInit#6 xAirValve');
    AssertEquals_BOOL(Expected := FALSE, Actual := fbOffAndInit.xWashPump, Message := 'OffAndInit#6 xWashPump');
    AssertEquals_BOOL(Expected := FALSE, Actual := fbOffAndInit.xInletValve, Message := 'OffAndInit#6 xInletValve');
    AssertEquals_BOOL(Expected := TRUE, Actual := fbOffAndInit.xWashActive, Message := 'OffAndInit#6 xWashActive');
    AssertEquals_BOOL(Expected := FALSE, Actual := fbOffAndInit.xValvesBusy, Message := 'OffAndInit#6 xValvesBusy');
    AssertEquals_INT(Expected := 1, Actual := fbOffAndInit.iWashCount, Message := 'OffAndInit#6 iWashCount');

    // #7, t = 600 мс — пуск: Drain, промывка №2
    GVL_S7Clock.tSimNow := T#600MS;
    fbOffAndInit.INIT_SQ := FALSE;
    fbOffAndInit.xStart := TRUE;
    fbOffAndInit();
    AssertEquals_BOOL(Expected := FALSE, Actual := fbOffAndInit.ERR_FLT, Message := 'OffAndInit#7 ERR_FLT');
    AssertEquals_BOOL(Expected := FALSE, Actual := fbOffAndInit.xReady, Message := 'OffAndInit#7 xReady');
    AssertEquals_BOOL(Expected := TRUE, Actual := fbOffAndInit.xDrainValve, Message := 'OffAndInit#7 xDrainValve');
    AssertEquals_BOOL(Expected := FALSE, Actual := fbOffAndInit.xBlower, Message := 'OffAndInit#7 xBlower');
    AssertEquals_BOOL(Expected := FALSE, Actual := fbOffAndInit.xAirValve, Message := 'OffAndInit#7 xAirValve');
    AssertEquals_BOOL(Expected := FALSE, Actual := fbOffAndInit.xWashPump, Message := 'OffAndInit#7 xWashPump');
    AssertEquals_BOOL(Expected := FALSE, Actual := fbOffAndInit.xInletValve, Message := 'OffAndInit#7 xInletValve');
    AssertEquals_BOOL(Expected := TRUE, Actual := fbOffAndInit.xWashActive, Message := 'OffAndInit#7 xWashActive');
    AssertEquals_BOOL(Expected := TRUE, Actual := fbOffAndInit.xValvesBusy, Message := 'OffAndInit#7 xValvesBusy');
    AssertEquals_INT(Expected := 2, Actual := fbOffAndInit.iWashCount, Message := 'OffAndInit#7 iWashCount');

    GVL_S7Clock.xSimulation := FALSE;
END_IF
coUnit.TEST_FINISHED();

(* ---- ShortWash.method.impl.st ---- *)
// AUTO-GENERATED — не редактировать: scenarios/lang/FB_BackwashGraph.csv, сценарий ShortWash
coUnit.TEST('ShortWash');
IF NOT xShortWashDone THEN
    xShortWashDone := TRUE;
    GVL_S7Clock.xSimulation := TRUE;

    // #1, t = 0 мс — первый вызов: начальный шаг Idle
    GVL_S7Clock.tSimNow := T#0MS;
    fbShortWash.OFF_SQ := FALSE;
    fbShortWash.INIT_SQ := FALSE;
    fbShortWash.ACK_EF := FALSE;
    fbShortWash.xStart := FALSE;
    fbShortWash.xLevelLow := FALSE;
    fbShortWash.xLevelHigh := FALSE;
    fbShortWash.xShortWash := FALSE;
    fbShortWash.xPumpOk := TRUE;
    fbShortWash.xValveFault := FALSE;
    fbShortWash();
    AssertEquals_BOOL(Expected := FALSE, Actual := fbShortWash.ERR_FLT, Message := 'ShortWash#1 ERR_FLT');
    AssertEquals_BOOL(Expected := TRUE, Actual := fbShortWash.xReady, Message := 'ShortWash#1 xReady');
    AssertEquals_BOOL(Expected := FALSE, Actual := fbShortWash.xDrainValve, Message := 'ShortWash#1 xDrainValve');
    AssertEquals_BOOL(Expected := FALSE, Actual := fbShortWash.xBlower, Message := 'ShortWash#1 xBlower');
    AssertEquals_BOOL(Expected := FALSE, Actual := fbShortWash.xAirValve, Message := 'ShortWash#1 xAirValve');
    AssertEquals_BOOL(Expected := FALSE, Actual := fbShortWash.xWashPump, Message := 'ShortWash#1 xWashPump');
    AssertEquals_BOOL(Expected := FALSE, Actual := fbShortWash.xInletValve, Message := 'ShortWash#1 xInletValve');
    AssertEquals_BOOL(Expected := FALSE, Actual := fbShortWash.xWashActive, Message := 'ShortWash#1 xWashActive');
    AssertEquals_BOOL(Expected := FALSE, Actual := fbShortWash.xValvesBusy, Message := 'ShortWash#1 xValvesBusy');
    AssertEquals_INT(Expected := 0, Actual := fbShortWash.iWashCount, Message := 'ShortWash#1 iWashCount');

    // #2, t = 100 мс — T1 Start: Drain, промывка №1, слив открыт
    GVL_S7Clock.tSimNow := T#100MS;
    fbShortWash.xStart := TRUE;
    fbShortWash();
    AssertEquals_BOOL(Expected := FALSE, Actual := fbShortWash.ERR_FLT, Message := 'ShortWash#2 ERR_FLT');
    AssertEquals_BOOL(Expected := FALSE, Actual := fbShortWash.xReady, Message := 'ShortWash#2 xReady');
    AssertEquals_BOOL(Expected := TRUE, Actual := fbShortWash.xDrainValve, Message := 'ShortWash#2 xDrainValve');
    AssertEquals_BOOL(Expected := FALSE, Actual := fbShortWash.xBlower, Message := 'ShortWash#2 xBlower');
    AssertEquals_BOOL(Expected := FALSE, Actual := fbShortWash.xAirValve, Message := 'ShortWash#2 xAirValve');
    AssertEquals_BOOL(Expected := FALSE, Actual := fbShortWash.xWashPump, Message := 'ShortWash#2 xWashPump');
    AssertEquals_BOOL(Expected := FALSE, Actual := fbShortWash.xInletValve, Message := 'ShortWash#2 xInletValve');
    AssertEquals_BOOL(Expected := TRUE, Actual := fbShortWash.xWashActive, Message := 'ShortWash#2 xWashActive');
    AssertEquals_BOOL(Expected := TRUE, Actual := fbShortWash.xValvesBusy, Message := 'ShortWash#2 xValvesBusy');
    AssertEquals_INT(Expected := 1, Actual := fbShortWash.iWashCount, Message := 'ShortWash#2 iWashCount');

    // #3, t = 200 мс — слив
    GVL_S7Clock.tSimNow := T#200MS;
    fbShortWash.xStart := FALSE;
    fbShortWash();
    AssertEquals_BOOL(Expected := FALSE, Actual := fbShortWash.ERR_FLT, Message := 'ShortWash#3 ERR_FLT');
    AssertEquals_BOOL(Expected := FALSE, Actual := fbShortWash.xReady, Message := 'ShortWash#3 xReady');
    AssertEquals_BOOL(Expected := TRUE, Actual := fbShortWash.xDrainValve, Message := 'ShortWash#3 xDrainValve');
    AssertEquals_BOOL(Expected := FALSE, Actual := fbShortWash.xBlower, Message := 'ShortWash#3 xBlower');
    AssertEquals_BOOL(Expected := FALSE, Actual := fbShortWash.xAirValve, Message := 'ShortWash#3 xAirValve');
    AssertEquals_BOOL(Expected := FALSE, Actual := fbShortWash.xWashPump, Message := 'ShortWash#3 xWashPump');
    AssertEquals_BOOL(Expected := FALSE, Actual := fbShortWash.xInletValve, Message := 'ShortWash#3 xInletValve');
    AssertEquals_BOOL(Expected := TRUE, Actual := fbShortWash.xWashActive, Message := 'ShortWash#3 xWashActive');
    AssertEquals_BOOL(Expected := TRUE, Actual := fbShortWash.xValvesBusy, Message := 'ShortWash#3 xValvesBusy');
    AssertEquals_INT(Expected := 1, Actual := fbShortWash.iWashCount, Message := 'ShortWash#3 iWashCount');

    // #4, t = 1000 мс — T3 ShortWash: QuickRinse
    GVL_S7Clock.tSimNow := T#1000MS;
    fbShortWash.xLevelLow := TRUE;
    fbShortWash.xShortWash := TRUE;
    fbShortWash();
    AssertEquals_BOOL(Expected := FALSE, Actual := fbShortWash.ERR_FLT, Message := 'ShortWash#4 ERR_FLT');
    AssertEquals_BOOL(Expected := FALSE, Actual := fbShortWash.xReady, Message := 'ShortWash#4 xReady');
    AssertEquals_BOOL(Expected := FALSE, Actual := fbShortWash.xDrainValve, Message := 'ShortWash#4 xDrainValve');
    AssertEquals_BOOL(Expected := FALSE, Actual := fbShortWash.xBlower, Message := 'ShortWash#4 xBlower');
    AssertEquals_BOOL(Expected := FALSE, Actual := fbShortWash.xAirValve, Message := 'ShortWash#4 xAirValve');
    AssertEquals_BOOL(Expected := TRUE, Actual := fbShortWash.xWashPump, Message := 'ShortWash#4 xWashPump');
    AssertEquals_BOOL(Expected := FALSE, Actual := fbShortWash.xInletValve, Message := 'ShortWash#4 xInletValve');
    AssertEquals_BOOL(Expected := TRUE, Actual := fbShortWash.xWashActive, Message := 'ShortWash#4 xWashActive');
    AssertEquals_BOOL(Expected := FALSE, Actual := fbShortWash.xValvesBusy, Message := 'ShortWash#4 xValvesBusy');
    AssertEquals_INT(Expected := 1, Actual := fbShortWash.iWashCount, Message := 'ShortWash#4 iWashCount');

    // #5, t = 1100 мс — быстрая отмывка
    GVL_S7Clock.tSimNow := T#1100MS;
    fbShortWash.xLevelLow := FALSE;
    fbShortWash();
    AssertEquals_BOOL(Expected := FALSE, Actual := fbShortWash.ERR_FLT, Message := 'ShortWash#5 ERR_FLT');
    AssertEquals_BOOL(Expected := FALSE, Actual := fbShortWash.xReady, Message := 'ShortWash#5 xReady');
    AssertEquals_BOOL(Expected := FALSE, Actual := fbShortWash.xDrainValve, Message := 'ShortWash#5 xDrainValve');
    AssertEquals_BOOL(Expected := FALSE, Actual := fbShortWash.xBlower, Message := 'ShortWash#5 xBlower');
    AssertEquals_BOOL(Expected := FALSE, Actual := fbShortWash.xAirValve, Message := 'ShortWash#5 xAirValve');
    AssertEquals_BOOL(Expected := TRUE, Actual := fbShortWash.xWashPump, Message := 'ShortWash#5 xWashPump');
    AssertEquals_BOOL(Expected := FALSE, Actual := fbShortWash.xInletValve, Message := 'ShortWash#5 xInletValve');
    AssertEquals_BOOL(Expected := TRUE, Actual := fbShortWash.xWashActive, Message := 'ShortWash#5 xWashActive');
    AssertEquals_BOOL(Expected := FALSE, Actual := fbShortWash.xValvesBusy, Message := 'ShortWash#5 xValvesBusy');
    AssertEquals_INT(Expected := 1, Actual := fbShortWash.iWashCount, Message := 'ShortWash#5 iWashCount');

    // #6, t = 2000 мс — T5 QuickDone: Refill
    GVL_S7Clock.tSimNow := T#2000MS;
    fbShortWash.xLevelHigh := TRUE;
    fbShortWash();
    AssertEquals_BOOL(Expected := FALSE, Actual := fbShortWash.ERR_FLT, Message := 'ShortWash#6 ERR_FLT');
    AssertEquals_BOOL(Expected := FALSE, Actual := fbShortWash.xReady, Message := 'ShortWash#6 xReady');
    AssertEquals_BOOL(Expected := FALSE, Actual := fbShortWash.xDrainValve, Message := 'ShortWash#6 xDrainValve');
    AssertEquals_BOOL(Expected := FALSE, Actual := fbShortWash.xBlower, Message := 'ShortWash#6 xBlower');
    AssertEquals_BOOL(Expected := FALSE, Actual := fbShortWash.xAirValve, Message := 'ShortWash#6 xAirValve');
    AssertEquals_BOOL(Expected := FALSE, Actual := fbShortWash.xWashPump, Message := 'ShortWash#6 xWashPump');
    AssertEquals_BOOL(Expected := TRUE, Actual := fbShortWash.xInletValve, Message := 'ShortWash#6 xInletValve');
    AssertEquals_BOOL(Expected := FALSE, Actual := fbShortWash.xWashActive, Message := 'ShortWash#6 xWashActive');
    AssertEquals_BOOL(Expected := TRUE, Actual := fbShortWash.xValvesBusy, Message := 'ShortWash#6 xValvesBusy');
    AssertEquals_INT(Expected := 1, Actual := fbShortWash.iWashCount, Message := 'ShortWash#6 iWashCount');

    // #7, t = 2100 мс — T6 Full: прыжок к Idle
    GVL_S7Clock.tSimNow := T#2100MS;
    fbShortWash();
    AssertEquals_BOOL(Expected := FALSE, Actual := fbShortWash.ERR_FLT, Message := 'ShortWash#7 ERR_FLT');
    AssertEquals_BOOL(Expected := TRUE, Actual := fbShortWash.xReady, Message := 'ShortWash#7 xReady');
    AssertEquals_BOOL(Expected := FALSE, Actual := fbShortWash.xDrainValve, Message := 'ShortWash#7 xDrainValve');
    AssertEquals_BOOL(Expected := FALSE, Actual := fbShortWash.xBlower, Message := 'ShortWash#7 xBlower');
    AssertEquals_BOOL(Expected := FALSE, Actual := fbShortWash.xAirValve, Message := 'ShortWash#7 xAirValve');
    AssertEquals_BOOL(Expected := FALSE, Actual := fbShortWash.xWashPump, Message := 'ShortWash#7 xWashPump');
    AssertEquals_BOOL(Expected := FALSE, Actual := fbShortWash.xInletValve, Message := 'ShortWash#7 xInletValve');
    AssertEquals_BOOL(Expected := FALSE, Actual := fbShortWash.xWashActive, Message := 'ShortWash#7 xWashActive');
    AssertEquals_BOOL(Expected := FALSE, Actual := fbShortWash.xValvesBusy, Message := 'ShortWash#7 xValvesBusy');
    AssertEquals_INT(Expected := 1, Actual := fbShortWash.iWashCount, Message := 'ShortWash#7 iWashCount');

    // #8, t = 2200 мс — готов
    GVL_S7Clock.tSimNow := T#2200MS;
    fbShortWash.xLevelHigh := FALSE;
    fbShortWash.xShortWash := FALSE;
    fbShortWash();
    AssertEquals_BOOL(Expected := FALSE, Actual := fbShortWash.ERR_FLT, Message := 'ShortWash#8 ERR_FLT');
    AssertEquals_BOOL(Expected := TRUE, Actual := fbShortWash.xReady, Message := 'ShortWash#8 xReady');
    AssertEquals_BOOL(Expected := FALSE, Actual := fbShortWash.xDrainValve, Message := 'ShortWash#8 xDrainValve');
    AssertEquals_BOOL(Expected := FALSE, Actual := fbShortWash.xBlower, Message := 'ShortWash#8 xBlower');
    AssertEquals_BOOL(Expected := FALSE, Actual := fbShortWash.xAirValve, Message := 'ShortWash#8 xAirValve');
    AssertEquals_BOOL(Expected := FALSE, Actual := fbShortWash.xWashPump, Message := 'ShortWash#8 xWashPump');
    AssertEquals_BOOL(Expected := FALSE, Actual := fbShortWash.xInletValve, Message := 'ShortWash#8 xInletValve');
    AssertEquals_BOOL(Expected := FALSE, Actual := fbShortWash.xWashActive, Message := 'ShortWash#8 xWashActive');
    AssertEquals_BOOL(Expected := FALSE, Actual := fbShortWash.xValvesBusy, Message := 'ShortWash#8 xValvesBusy');
    AssertEquals_INT(Expected := 1, Actual := fbShortWash.iWashCount, Message := 'ShortWash#8 iWashCount');

    GVL_S7Clock.xSimulation := FALSE;
END_IF
coUnit.TEST_FINISHED();

(* ---- Supervision.method.impl.st ---- *)
// AUTO-GENERATED — не редактировать: scenarios/lang/FB_BackwashGraph.csv, сценарий Supervision
coUnit.TEST('Supervision');
IF NOT xSupervisionDone THEN
    xSupervisionDone := TRUE;
    GVL_S7Clock.xSimulation := TRUE;

    // #1, t = 0 мс — первый вызов: начальный шаг Idle
    GVL_S7Clock.tSimNow := T#0MS;
    fbSupervision.OFF_SQ := FALSE;
    fbSupervision.INIT_SQ := FALSE;
    fbSupervision.ACK_EF := FALSE;
    fbSupervision.xStart := FALSE;
    fbSupervision.xLevelLow := FALSE;
    fbSupervision.xLevelHigh := FALSE;
    fbSupervision.xShortWash := FALSE;
    fbSupervision.xPumpOk := TRUE;
    fbSupervision.xValveFault := FALSE;
    fbSupervision();
    AssertEquals_BOOL(Expected := FALSE, Actual := fbSupervision.ERR_FLT, Message := 'Supervision#1 ERR_FLT');
    AssertEquals_BOOL(Expected := TRUE, Actual := fbSupervision.xReady, Message := 'Supervision#1 xReady');
    AssertEquals_BOOL(Expected := FALSE, Actual := fbSupervision.xDrainValve, Message := 'Supervision#1 xDrainValve');
    AssertEquals_BOOL(Expected := FALSE, Actual := fbSupervision.xBlower, Message := 'Supervision#1 xBlower');
    AssertEquals_BOOL(Expected := FALSE, Actual := fbSupervision.xAirValve, Message := 'Supervision#1 xAirValve');
    AssertEquals_BOOL(Expected := FALSE, Actual := fbSupervision.xWashPump, Message := 'Supervision#1 xWashPump');
    AssertEquals_BOOL(Expected := FALSE, Actual := fbSupervision.xInletValve, Message := 'Supervision#1 xInletValve');
    AssertEquals_BOOL(Expected := FALSE, Actual := fbSupervision.xWashActive, Message := 'Supervision#1 xWashActive');
    AssertEquals_BOOL(Expected := FALSE, Actual := fbSupervision.xValvesBusy, Message := 'Supervision#1 xValvesBusy');
    AssertEquals_INT(Expected := 0, Actual := fbSupervision.iWashCount, Message := 'Supervision#1 iWashCount');

    // #2, t = 100 мс — T1 Start: Drain, промывка №1, слив открыт
    GVL_S7Clock.tSimNow := T#100MS;
    fbSupervision.xStart := TRUE;
    fbSupervision();
    AssertEquals_BOOL(Expected := FALSE, Actual := fbSupervision.ERR_FLT, Message := 'Supervision#2 ERR_FLT');
    AssertEquals_BOOL(Expected := FALSE, Actual := fbSupervision.xReady, Message := 'Supervision#2 xReady');
    AssertEquals_BOOL(Expected := TRUE, Actual := fbSupervision.xDrainValve, Message := 'Supervision#2 xDrainValve');
    AssertEquals_BOOL(Expected := FALSE, Actual := fbSupervision.xBlower, Message := 'Supervision#2 xBlower');
    AssertEquals_BOOL(Expected := FALSE, Actual := fbSupervision.xAirValve, Message := 'Supervision#2 xAirValve');
    AssertEquals_BOOL(Expected := FALSE, Actual := fbSupervision.xWashPump, Message := 'Supervision#2 xWashPump');
    AssertEquals_BOOL(Expected := FALSE, Actual := fbSupervision.xInletValve, Message := 'Supervision#2 xInletValve');
    AssertEquals_BOOL(Expected := TRUE, Actual := fbSupervision.xWashActive, Message := 'Supervision#2 xWashActive');
    AssertEquals_BOOL(Expected := TRUE, Actual := fbSupervision.xValvesBusy, Message := 'Supervision#2 xValvesBusy');
    AssertEquals_INT(Expected := 1, Actual := fbSupervision.iWashCount, Message := 'Supervision#2 iWashCount');

    // #3, t = 200 мс — слив
    GVL_S7Clock.tSimNow := T#200MS;
    fbSupervision.xStart := FALSE;
    fbSupervision();
    AssertEquals_BOOL(Expected := FALSE, Actual := fbSupervision.ERR_FLT, Message := 'Supervision#3 ERR_FLT');
    AssertEquals_BOOL(Expected := FALSE, Actual := fbSupervision.xReady, Message := 'Supervision#3 xReady');
    AssertEquals_BOOL(Expected := TRUE, Actual := fbSupervision.xDrainValve, Message := 'Supervision#3 xDrainValve');
    AssertEquals_BOOL(Expected := FALSE, Actual := fbSupervision.xBlower, Message := 'Supervision#3 xBlower');
    AssertEquals_BOOL(Expected := FALSE, Actual := fbSupervision.xAirValve, Message := 'Supervision#3 xAirValve');
    AssertEquals_BOOL(Expected := FALSE, Actual := fbSupervision.xWashPump, Message := 'Supervision#3 xWashPump');
    AssertEquals_BOOL(Expected := FALSE, Actual := fbSupervision.xInletValve, Message := 'Supervision#3 xInletValve');
    AssertEquals_BOOL(Expected := TRUE, Actual := fbSupervision.xWashActive, Message := 'Supervision#3 xWashActive');
    AssertEquals_BOOL(Expected := TRUE, Actual := fbSupervision.xValvesBusy, Message := 'Supervision#3 xValvesBusy');
    AssertEquals_INT(Expected := 1, Actual := fbSupervision.iWashCount, Message := 'Supervision#3 iWashCount');

    // #4, t = 500 мс — неисправность задвижки: ERR_FLT
    GVL_S7Clock.tSimNow := T#500MS;
    fbSupervision.xValveFault := TRUE;
    fbSupervision();
    AssertEquals_BOOL(Expected := TRUE, Actual := fbSupervision.ERR_FLT, Message := 'Supervision#4 ERR_FLT');
    AssertEquals_BOOL(Expected := FALSE, Actual := fbSupervision.xReady, Message := 'Supervision#4 xReady');
    AssertEquals_BOOL(Expected := TRUE, Actual := fbSupervision.xDrainValve, Message := 'Supervision#4 xDrainValve');
    AssertEquals_BOOL(Expected := FALSE, Actual := fbSupervision.xBlower, Message := 'Supervision#4 xBlower');
    AssertEquals_BOOL(Expected := FALSE, Actual := fbSupervision.xAirValve, Message := 'Supervision#4 xAirValve');
    AssertEquals_BOOL(Expected := FALSE, Actual := fbSupervision.xWashPump, Message := 'Supervision#4 xWashPump');
    AssertEquals_BOOL(Expected := FALSE, Actual := fbSupervision.xInletValve, Message := 'Supervision#4 xInletValve');
    AssertEquals_BOOL(Expected := TRUE, Actual := fbSupervision.xWashActive, Message := 'Supervision#4 xWashActive');
    AssertEquals_BOOL(Expected := TRUE, Actual := fbSupervision.xValvesBusy, Message := 'Supervision#4 xValvesBusy');
    AssertEquals_INT(Expected := 1, Actual := fbSupervision.iWashCount, Message := 'Supervision#4 iWashCount');

    // #5, t = 600 мс — уровень низкий, но переход заблокирован ошибкой
    GVL_S7Clock.tSimNow := T#600MS;
    fbSupervision.xLevelLow := TRUE;
    fbSupervision();
    AssertEquals_BOOL(Expected := TRUE, Actual := fbSupervision.ERR_FLT, Message := 'Supervision#5 ERR_FLT');
    AssertEquals_BOOL(Expected := FALSE, Actual := fbSupervision.xReady, Message := 'Supervision#5 xReady');
    AssertEquals_BOOL(Expected := TRUE, Actual := fbSupervision.xDrainValve, Message := 'Supervision#5 xDrainValve');
    AssertEquals_BOOL(Expected := FALSE, Actual := fbSupervision.xBlower, Message := 'Supervision#5 xBlower');
    AssertEquals_BOOL(Expected := FALSE, Actual := fbSupervision.xAirValve, Message := 'Supervision#5 xAirValve');
    AssertEquals_BOOL(Expected := FALSE, Actual := fbSupervision.xWashPump, Message := 'Supervision#5 xWashPump');
    AssertEquals_BOOL(Expected := FALSE, Actual := fbSupervision.xInletValve, Message := 'Supervision#5 xInletValve');
    AssertEquals_BOOL(Expected := TRUE, Actual := fbSupervision.xWashActive, Message := 'Supervision#5 xWashActive');
    AssertEquals_BOOL(Expected := TRUE, Actual := fbSupervision.xValvesBusy, Message := 'Supervision#5 xValvesBusy');
    AssertEquals_INT(Expected := 1, Actual := fbSupervision.iWashCount, Message := 'Supervision#5 iWashCount');

    // #6, t = 700 мс — квитирование при неисправности: ошибка сразу снова
    GVL_S7Clock.tSimNow := T#700MS;
    fbSupervision.ACK_EF := TRUE;
    fbSupervision.xLevelLow := FALSE;
    fbSupervision();
    AssertEquals_BOOL(Expected := TRUE, Actual := fbSupervision.ERR_FLT, Message := 'Supervision#6 ERR_FLT');
    AssertEquals_BOOL(Expected := FALSE, Actual := fbSupervision.xReady, Message := 'Supervision#6 xReady');
    AssertEquals_BOOL(Expected := TRUE, Actual := fbSupervision.xDrainValve, Message := 'Supervision#6 xDrainValve');
    AssertEquals_BOOL(Expected := FALSE, Actual := fbSupervision.xBlower, Message := 'Supervision#6 xBlower');
    AssertEquals_BOOL(Expected := FALSE, Actual := fbSupervision.xAirValve, Message := 'Supervision#6 xAirValve');
    AssertEquals_BOOL(Expected := FALSE, Actual := fbSupervision.xWashPump, Message := 'Supervision#6 xWashPump');
    AssertEquals_BOOL(Expected := FALSE, Actual := fbSupervision.xInletValve, Message := 'Supervision#6 xInletValve');
    AssertEquals_BOOL(Expected := TRUE, Actual := fbSupervision.xWashActive, Message := 'Supervision#6 xWashActive');
    AssertEquals_BOOL(Expected := TRUE, Actual := fbSupervision.xValvesBusy, Message := 'Supervision#6 xValvesBusy');
    AssertEquals_INT(Expected := 1, Actual := fbSupervision.iWashCount, Message := 'Supervision#6 iWashCount');

    // #7, t = 800 мс — неисправность ушла, ошибка держится
    GVL_S7Clock.tSimNow := T#800MS;
    fbSupervision.ACK_EF := FALSE;
    fbSupervision.xValveFault := FALSE;
    fbSupervision();
    AssertEquals_BOOL(Expected := TRUE, Actual := fbSupervision.ERR_FLT, Message := 'Supervision#7 ERR_FLT');
    AssertEquals_BOOL(Expected := FALSE, Actual := fbSupervision.xReady, Message := 'Supervision#7 xReady');
    AssertEquals_BOOL(Expected := TRUE, Actual := fbSupervision.xDrainValve, Message := 'Supervision#7 xDrainValve');
    AssertEquals_BOOL(Expected := FALSE, Actual := fbSupervision.xBlower, Message := 'Supervision#7 xBlower');
    AssertEquals_BOOL(Expected := FALSE, Actual := fbSupervision.xAirValve, Message := 'Supervision#7 xAirValve');
    AssertEquals_BOOL(Expected := FALSE, Actual := fbSupervision.xWashPump, Message := 'Supervision#7 xWashPump');
    AssertEquals_BOOL(Expected := FALSE, Actual := fbSupervision.xInletValve, Message := 'Supervision#7 xInletValve');
    AssertEquals_BOOL(Expected := TRUE, Actual := fbSupervision.xWashActive, Message := 'Supervision#7 xWashActive');
    AssertEquals_BOOL(Expected := TRUE, Actual := fbSupervision.xValvesBusy, Message := 'Supervision#7 xValvesBusy');
    AssertEquals_INT(Expected := 1, Actual := fbSupervision.iWashCount, Message := 'Supervision#7 iWashCount');

    // #8, t = 900 мс — квитирование: ошибка снята
    GVL_S7Clock.tSimNow := T#900MS;
    fbSupervision.ACK_EF := TRUE;
    fbSupervision();
    AssertEquals_BOOL(Expected := FALSE, Actual := fbSupervision.ERR_FLT, Message := 'Supervision#8 ERR_FLT');
    AssertEquals_BOOL(Expected := FALSE, Actual := fbSupervision.xReady, Message := 'Supervision#8 xReady');
    AssertEquals_BOOL(Expected := TRUE, Actual := fbSupervision.xDrainValve, Message := 'Supervision#8 xDrainValve');
    AssertEquals_BOOL(Expected := FALSE, Actual := fbSupervision.xBlower, Message := 'Supervision#8 xBlower');
    AssertEquals_BOOL(Expected := FALSE, Actual := fbSupervision.xAirValve, Message := 'Supervision#8 xAirValve');
    AssertEquals_BOOL(Expected := FALSE, Actual := fbSupervision.xWashPump, Message := 'Supervision#8 xWashPump');
    AssertEquals_BOOL(Expected := FALSE, Actual := fbSupervision.xInletValve, Message := 'Supervision#8 xInletValve');
    AssertEquals_BOOL(Expected := TRUE, Actual := fbSupervision.xWashActive, Message := 'Supervision#8 xWashActive');
    AssertEquals_BOOL(Expected := TRUE, Actual := fbSupervision.xValvesBusy, Message := 'Supervision#8 xValvesBusy');
    AssertEquals_INT(Expected := 1, Actual := fbSupervision.iWashCount, Message := 'Supervision#8 iWashCount');

    // #9, t = 1000 мс — T2 LongWash: Air и Rinse
    GVL_S7Clock.tSimNow := T#1000MS;
    fbSupervision.ACK_EF := FALSE;
    fbSupervision.xLevelLow := TRUE;
    fbSupervision();
    AssertEquals_BOOL(Expected := FALSE, Actual := fbSupervision.ERR_FLT, Message := 'Supervision#9 ERR_FLT');
    AssertEquals_BOOL(Expected := FALSE, Actual := fbSupervision.xReady, Message := 'Supervision#9 xReady');
    AssertEquals_BOOL(Expected := FALSE, Actual := fbSupervision.xDrainValve, Message := 'Supervision#9 xDrainValve');
    AssertEquals_BOOL(Expected := TRUE, Actual := fbSupervision.xBlower, Message := 'Supervision#9 xBlower');
    AssertEquals_BOOL(Expected := FALSE, Actual := fbSupervision.xAirValve, Message := 'Supervision#9 xAirValve');
    AssertEquals_BOOL(Expected := TRUE, Actual := fbSupervision.xWashPump, Message := 'Supervision#9 xWashPump');
    AssertEquals_BOOL(Expected := FALSE, Actual := fbSupervision.xInletValve, Message := 'Supervision#9 xInletValve');
    AssertEquals_BOOL(Expected := TRUE, Actual := fbSupervision.xWashActive, Message := 'Supervision#9 xWashActive');
    AssertEquals_BOOL(Expected := FALSE, Actual := fbSupervision.xValvesBusy, Message := 'Supervision#9 xValvesBusy');
    AssertEquals_INT(Expected := 1, Actual := fbSupervision.iWashCount, Message := 'Supervision#9 iWashCount');

    GVL_S7Clock.xSimulation := FALSE;
END_IF
coUnit.TEST_FINISHED();
